(* IEC 61131-3 sources: rusty/tests/lit/multi/real_remainder_shared, 2 files *)

(* ---- main.st ---- *)
FUNCTION main : DINT
    printf('REAL: %.2f$N', REAL_TO_LREAL(remainderReal(7.5, 2.0)));
    printf('LREAL: %.2f$N', remainderLreal(-7.5, 2.0));
END_FUNCTION

(* ---- remainder.st ---- *)
FUNCTION remainderReal : REAL
VAR_INPUT
    value, range : REAL;
END_VAR
    remainderReal := value MOD range;
END_FUNCTION

FUNCTION remainderLreal : LREAL
VAR_INPUT
    value, range : LREAL;
END_VAR
    remainderLreal := value MOD range;
END_FUNCTION
